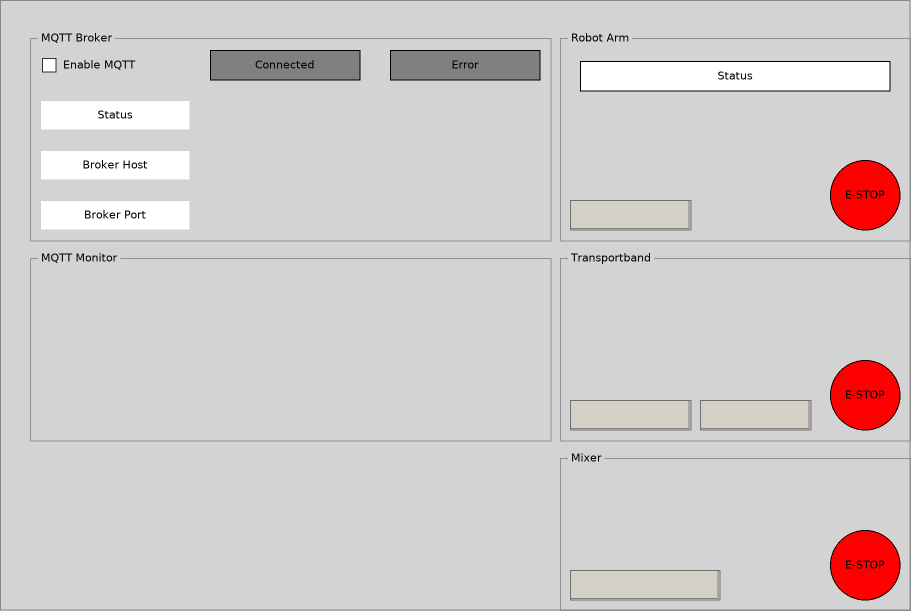
VISUALIZATION PannenkoekenDashboard  // 911x611
    GroupBox (30,30 521x211), "MQTT Broker"
        Checkbox (10,20 150x30), "Enable MQTT"
        Rectangle (360,20 150x30), "Error"
        Rectangle (180,20 150x30), "Connected"
        Textfield (10,70 150x30), "Status"
        Textfield (10,120 150x30), "Broker Host"
        Textfield (10,170 150x30), "Broker Port"
    GroupBox (30,250 521x191), "MQTT Monitor"
    GroupBox (560,30 351x211), "Robot Arm"
        Rectangle (20,31 310x30), "Status"
        Ellipse (270,130 70x70), "E-STOP"
        Button (10,170 121x30)
    GroupBox (560,250 351x191), "Transportband"
        Ellipse (270,110 70x70), "E-STOP"
        Button (10,150 121x30)
        Button (140,150 111x30)
    GroupBox (560,450 351x161), "Mixer"
        Ellipse (270,80 70x70), "E-STOP"
        Button (10,120 150x30)
END_VISUALIZATION

(* stored: Version 1.1.0.1, ProductVersion 3.1.4024.15
   Visu PannenkoekenDashboard: Id {747fc4aa-41f4-4f69-b086-b41493138125} *)
